  # add a "skill" to the robots skillset the control system will send a string with the ls_item and action and here we will look if we have a matching skill to execute
  # the item_modell defines the patterns which have to be used by the robot on multiple racks and or multiple samples in a rackpattern
  # inner pattern is always dependung on the object that has to be moved and the outer pattern is the pattern for the containers where the objects are stored in.
  # if racks have to be handled it is also an inner pattern cause the object to handle is the rack itself
  # create_item(id=0, ls_item="default", frame=p[0,0,0,0,0,0], actionlist=create_action_list([]), item_model=create_item_model(), lm_id=0, description="default")
  # create_item_model(inner=create_pattern(), outer=create_pattern(), description="default")
  # ITEM_MAP.append(create_item(id=1, ls_item="Home", frame=F1_uLM_Home, actionlist=[ActionManipulator.MOVE_TO], description="uLM Move To Home"))
  # ITEM_MAP.append(create_item(id=2, ls_item="InputStation", frame=F2_uLM_Input, actionlist=[ActionManipulator.PICK, ActionManipulator.PLACE], item_model=create_item_model(inner=Patterns.INPUT), description="uLM Pick and Place samples from Input"))
  # ITEM_MAP.append(create_item(id=3, ls_item="InputCapture", frame=F3_Cap_Input, actionlist=[ActionCamera.INSPECT, ActionManipulator.MOVE_TO], description="uLM Inspect samples from Input and Move To Capture Position"))
  # ITEM_MAP.append(create_item(id=4, ls_item="Bin", frame=F4_uLM_Bin, actionlist=[ActionManipulator.PLACE], description="uLM Place Cap to Bin"))
  # ITEM_MAP.append(create_item(id=5, ls_item="StationaryGripper", frame=F5_uLM_Gripper, actionlist=[ActionManipulator.PICK, ActionManipulator.PLACE, ActionManipulator.DECAP, ActionManipulator.MOVE_TO, ActionManipulator.GRASP, ActionManipulator.RELEASE], description=" uLM stationary gripper"))
  # ITEM_MAP.append(create_item(id=6, ls_item="CobasRack", frame=F6_uLM_Cobas_R, actionlist=[ActionManipulator.PICK, ActionManipulator.PLACE], item_model=create_item_model(outer=Patterns.COBAS_MAGAZINE), description="uLM Cobas Racks Pick and Place"))
  # ITEM_MAP.append(create_item(id=7, ls_item="CobasMagazine", frame=F7_uLM_Coba_Mag, actionlist=[ActionManipulator.PICK, ActionManipulator.PLACE], item_model=create_item_model(inner=Patterns.COBAS, outer=Patterns.COBAS_MAGAZINE), description="uLM Cobas Magazine Samples Pick and Place"))
  # ITEM_MAP.append(create_item(id=8, ls_item="DetectCobasRacks", frame=F8_Cap_Cobas_LM, actionlist=[ActionCamera.DETECT_OBJECTS, ActionManipulator.MOVE_TO], lm_id=2, description="uLM Cobas Rack Detection and Move To Capture"))
  # ITEM_MAP.append(create_item(id=9, ls_item="TaraMagazine", frame=F9_uLM_Tara, actionlist=[ActionManipulator.PICK, ActionManipulator.PLACE], item_model=create_item_model(inner=Patterns.TARA), description="uLM Centrifuge Tara Pick and Place"))
  # ITEM_MAP.append(create_item(id=10, ls_item="CentrifugeCapture", frame=F10_Cap_CF, actionlist=[ActionManipulator.MOVE_TO, ActionCamera.DETECT], lm_id=1, description="Centrifuge Device Move to Capture Pos and Detect Landmarks"))
  # ITEM_MAP.append(create_item(id=11, ls_item="Centrifuge", frame=F11_CF_PiPl, actionlist=[ActionManipulator.PICK, ActionManipulator.PLACE], description="Centrifuge Device Rack Pick and Place"))
  # ITEM_MAP.append(create_item(id=12, ls_item="CentrifugeMagazine", frame=F12_uLM_CF_Mag, actionlist=[ActionManipulator.PICK, ActionManipulator.PLACE], item_model=create_item_model(inner=Patterns.CENTRIFUGE, outer=Patterns.CENTRIFUGE_MAGAZINE), description=" uLM Centrifuge Magazin Pick and Place"))
  # ITEM_MAP.append(create_item(id=13, ls_item="CentrifugeRack", frame=F13_uLM_CF_R, actionlist=[ActionManipulator.PICK, ActionManipulator.PLACE], item_model=create_item_model(outer=Patterns.CENTRIFUGE_MAGAZINE), description="uLM Centrifuge Magazin Pick and Place Racks"))
  # ITEM_MAP.append(create_item(id=14, ls_item="DailyArchive", frame=F14_uLM_Archive, actionlist=[ActionManipulator.PICK, ActionManipulator.PLACE], item_model=create_item_model(inner=Patterns.ARCHIVE), description="uLM Pick and Place samples from Archive Rack"))
  # ITEM_MAP.append(create_item(id=15, ls_item="NokRack", frame=F15_uLM_Nok, actionlist=[ActionManipulator.PICK, ActionManipulator.PLACE], item_model=create_item_model(inner=Patterns.NOK), description="uLM Pick and Place samples from Nok Rack"))
  # ITEM_MAP.append(create_item(id=16, ls_item="CobasInput", frame=F16_Cobas_Input, actionlist=[ActionManipulator.PLACE], description="uLM Place Cobasrack in Cobas Device"))
  # ITEM_MAP.append(create_item(id=17, ls_item="CobasInputCapture", frame=F17_Cobas_Cap, actionlist=[ActionCamera.DETECT, ActionManipulator.MOVE_TO], lm_id=3, description="uLM Place Cobasrack in Cobas Device"))
  # ITEM_MAP.append(create_item(id=18, ls_item="XN550Input", frame=F18_XN550_Input, actionlist=[ActionManipulator.PICK, ActionManipulator.PLACE], item_model=create_item_model(inner=Patterns.SYSMEX_XN550, outer=Patterns.DRAWER_XN550), lm_id=4, description="uLM Pick and Place Samples in or out of XN550 Racks"))
  # ITEM_MAP.append(create_item(id=19, ls_item="XN550Capture", frame=F19_XN550_Cap, actionlist=[ActionCamera.DETECT, ActionManipulator.MOVE_TO], lm_id=4, description="uLM Move To and Capture LM XN550"))
  # ITEM_MAP.append(create_item(id=20, ls_item="XN550Drawer", frame=F20_XN550_Draw, actionlist=[ActionManipulator.DRAWER_OPEN, ActionManipulator.DRAWER_CLOSE], item_model=create_item_model(inner=Patterns.DRAWER_XN550), lm_id=4, description="uLM Open and close Drawer XN550"))
  # ITEM_MAP.append(create_item(id=21, ls_item="XN550Button", frame=F21_XN550_Btn, actionlist=[ActionManipulator.PUSH], lm_id=4, description="uLM Push XN550 Button"))
  # ITEM_MAP.append(create_item(id=22, ls_item="AMR", frame=p[0,0,0,0,0,0], actionlist=[ActionAMR.READ, ActionAMR.LOAD_MISSION, ActionAMR.START_MISSION, ActionAMR.NAVIGATE, ActionAMR.ACKNOWLEDGE], description="all AMR actions"))



  # ITEM_MAP.append(create_item(id=31, ls_item="TestLM", frame=TestLM, actionlist=[ActionManipulator.PICK, ActionManipulator.PLACE], item_model=create_item_model(inner=Rack.SYSMEX_CS2500), lm_id=5, description="LM Test"))
  # Fills the Vision Config List with Projectrelated Data
  # workspaceid and skillid are highly robominds related so probably will not stay like this in the future
  # sample detection: dx and dy are used to calculate the positions in a rack and given by the offset which will be applied in order to assign the sample to a place in the rack
  # create_vision_config(workspace_id="", skill_id="", item_id=-1, capture_pos=p[0,0,0,0,0,0], dx=0, dy=0, target_origin=p[0,0,0,0,0,0], selector="default", description="default")
  # VISION_CONFIG_MAP.append(create_vision_config(workspace_id="96017791-f581-4e9e-93da-6951695fccc8", skill_id="8885cfe1-6784-4293-bd26-52ebdc67bf95", capture_pos=F10_Cap_CF, target_origin=p[0,0,0,0,0,0], item_id=11, description="LM Detect CF"))
  # VISION_CONFIG_MAP.append(create_vision_config(workspace_id="96017791-f581-4e9e-93da-6951695fccc8", skill_id="8885cfe1-6784-4293-bd26-52ebdc67bf95", capture_pos=F8_Cap_Cobas_LM, target_origin=p[0,0,0,0,0,0], item_id=8, description="LM Detect Cobas Racks"))
  # VISION_CONFIG_MAP.append(create_vision_config(workspace_id="8f0ad01c-dc36-4fdd-b295-0b6b4a38b89a", skill_id="afdc9e13-ea83-40d6-a805-bb041453d2e5", capture_pos=F3_Cap_Input, target_origin=F2_uLM_Input, item_id=3, description="Lab Solution Input Capture"))
  # VISION_CONFIG_MAP.append(create_vision_config(workspace_id="96017791-f581-4e9e-93da-6951695fccc8", skill_id="8885cfe1-6784-4293-bd26-52ebdc67bf95", capture_pos=F19_XN550_Cap, target_origin=F18_XN550_Input, item_id=18, description="Input XN550"))
  # VISION_CONFIG_MAP.append(create_vision_config(workspace_id="96017791-f581-4e9e-93da-6951695fccc8", skill_id="8885cfe1-6784-4293-bd26-52ebdc67bf95", capture_pos=F19_XN550_Cap, target_origin=POS_Z, item_id=19, description="LM Detect XN550F"))
  # VISION_CONFIG_MAP.append(create_vision_config(workspace_id="96017791-f581-4e9e-93da-6951695fccc8", skill_id="8885cfe1-6784-4293-bd26-52ebdc67bf95", capture_pos=F10_Cap_CF, target_origin=POS_Z, item_id=10, description="LM Detect CF"))
  # VISION_CONFIG_MAP.append(create_vision_config(workspace_id="96017791-f581-4e9e-93da-6951695fccc8", skill_id="8885cfe1-6784-4293-bd26-52ebdc67bf95", capture_pos=F19_XN550_Cap, target_origin=F20_XN550_Draw, item_id=20, description="Drawer XN550"))
  # VISION_CONFIG_MAP.append(create_vision_config(workspace_id="96017791-f581-4e9e-93da-6951695fccc8", skill_id="8885cfe1-6784-4293-bd26-52ebdc67bf95", capture_pos=F19_XN550_Cap, target_origin=F21_XN550_Btn, item_id=21, description="Button XN550"))
  # VISION_CONFIG_MAP.append(create_vision_config(workspace_id="96017791-f581-4e9e-93da-6951695fccc8", skill_id="8885cfe1-6784-4293-bd26-52ebdc67bf95", capture_pos=TestLMCap, target_origin=p[0,0,0,0,0,0], item_id=30, description="Button XN550"))
  # VISION_CONFIG_MAP.append(create_vision_config(workspace_id="96017791-f581-4e9e-93da-6951695fccc8", skill_id="8885cfe1-6784-4293-bd26-52ebdc67bf95", capture_pos=TestLMCap, target_origin=TestLM, item_id=31, description="Button XN550"))

  # VISION_CONFIG_MAP.append(create_vision_config(workspace_id="96017791-f581-4e9e-93da-6951695fccc8", skill_id="8885cfe1-6784-4293-bd26-52ebdc67bf95", target_origin=p[0,0,0,0,0,0], item_id=11, description="LM Detect CF"))
  # VISION_CONFIG_MAP.append(create_vision_config(workspace_id="96017791-f581-4e9e-93da-6951695fccc8", skill_id="8885cfe1-6784-4293-bd26-52ebdc67bf95", target_origin=p[0,0,0,0,0,0], item_id=8, description="LM Detect Cobas Racks"))
  # VISION_CONFIG_MAP.append(create_vision_config(workspace_id="8f0ad01c-dc36-4fdd-b295-0b6b4a38b89a", skill_id="afdc9e13-ea83-40d6-a805-bb041453d2e5", target_origin=F2_uLM_Input, item_id=3, description="Lab Solution Input Capture"))
  # VISION_CONFIG_MAP.append(create_vision_config(workspace_id="96017791-f581-4e9e-93da-6951695fccc8", skill_id="8885cfe1-6784-4293-bd26-52ebdc67bf95", target_origin=F18_XN550_Input, item_id=18, description="Input XN550"))
  # VISION_CONFIG_MAP.append(create_vision_config(workspace_id="96017791-f581-4e9e-93da-6951695fccc8", skill_id="8885cfe1-6784-4293-bd26-52ebdc67bf95", target_origin=POS_Z, item_id=19, description="LM Detect XN550F"))
  # VISION_CONFIG_MAP.append(create_vision_config(workspace_id="96017791-f581-4e9e-93da-6951695fccc8", skill_id="8885cfe1-6784-4293-bd26-52ebdc67bf95", target_origin=POS_Z, item_id=10, description="LM Detect CF"))
  # VISION_CONFIG_MAP.append(create_vision_config(workspace_id="96017791-f581-4e9e-93da-6951695fccc8", skill_id="8885cfe1-6784-4293-bd26-52ebdc67bf95", target_origin=F20_XN550_Draw, item_id=20, description="Drawer XN550"))
  # VISION_CONFIG_MAP.append(create_vision_config(workspace_id="96017791-f581-4e9e-93da-6951695fccc8", skill_id="8885cfe1-6784-4293-bd26-52ebdc67bf95", target_origin=F21_XN550_Btn, item_id=21, description="Button XN550"))
  # VISION_CONFIG_MAP.append(create_vision_config(workspace_id="96017791-f581-4e9e-93da-6951695fccc8", skill_id="8885cfe1-6784-4293-bd26-52ebdc67bf95", target_origin=p[0,0,0,0,0,0], item_id=30, description="Button XN550"))
  # VISION_CONFIG_MAP.append(create_vision_config(workspace_id="96017791-f581-4e9e-93da-6951695fccc8", skill_id="8885cfe1-6784-4293-bd26-52ebdc67bf95", target_origin=TestLM, item_id=31, description="Button XN550"))

  # local inputrack = find_pattern_by_name("INPUT")
  # INSPECT_CONFIG_MAP.append(create_inspect_config(item_id=3, dx=inputrack.pattern_width[0]/(inputrack.pattern_size[0]-1), dy=inputrack.pattern_width[1]/(inputrack.pattern_size[1]-1), rack_size=inputrack.pattern_size , description="Input Capture"))
  # # Fills the Landmark List with Projectrelated Data
  # # create_landmark(lm_id=0, marker_id=-1, marker_size=0.1, marker_type="aruco_7x7", capture_pos=p[0,0,0,0,0,0], init_frame=p[0,0,0,0,0,0], search_offset=[0,0,0], actual_frame=p[0,0,0,0,0,0], description="")
  # LANDMARK_MAP.append(create_landmark(lm_id=1, marker_id=3, marker_size=0.1, marker_type="aruco_7x7", capture_pos = F10_Cap_CF, init_frame=p[-0.617789, -0.065471, 0.07918, 0.020983, -0.012695, 1.512066], search_offset=[0.15, 0.15, 0.1], actual_frame=p[-0.617789, -0.065471, 0.07918, 0.020983, -0.012695, 1.512066], description="LM CF Lid"))
  # LANDMARK_MAP.append(create_landmark(lm_id=2, marker_id=-1, marker_size=0.0085, marker_type="aruco_4x4", capture_pos = F8_Cap_Cobas_LM, init_frame=p[0,0,0,0,0,0], search_offset=[0.15, 0.15, 0.1], actual_frame=POS_Z, description="LM Cobas Rack Detection"))
  # LANDMARK_MAP.append(create_landmark(lm_id=3, marker_id=0, marker_size=0.1, marker_type="aruco_7x7", capture_pos = F17_Cobas_Cap, init_frame=p[-0.667,-0.194,0.100,0,0,0], search_offset=[0.15, 0.15, 0.1], actual_frame=POS_Z, description="LM Cobas Cap"))
  # LANDMARK_MAP.append(create_landmark(lm_id=4, marker_id=4, marker_size=0.1, marker_type="aruco_7x7", capture_pos = F19_XN550_Cap, init_frame=p[0.124,-0.976,0.355,-0.008,0.025,3.131], search_offset=[0.15, 0.15, 0.1], actual_frame=p[0,0,0,0,0,0], description="LM XN550 Cap"))
  # LANDMARK_MAP.append(create_landmark(lm_id=5, marker_id=0, marker_size=0.1, marker_type="aruco_7x7", capture_pos = TestLMCap, init_frame=p[-0.49,-0.144,0.092,0,-0.008,0.001], search_offset=[0.15, 0.15, 0.1], actual_frame=POS_Z, description="LM Test"))
  # # Configuration of all movement related parameters
  # # create_movement(id=0, hh_approach=POS_Z, h_approach=POS_Z, approach=POS_Z, h_target=POS_Z, target=POS_Z, retract=POS_Z, h_retract=POS_Z, hh_retract=POS_Z, h_frame=POS_Z, frame=POS_Z, speed=1, acceleration=1, description="default")
  # MOVEMENT_MAP.append(create_movement(description="TestLMCap", frame=TestLMCap, actionlist=[ActionManipulator.MOVE_TO]))
  # MOVEMENT_MAP.append(create_movement(description="TestLM", frame=TestLM, actionlist=[ActionManipulator.PICK,ActionManipulator.PLACE],
  #         approach=p[0,0,0.1,0,0,0],
  #         retract=p[0,0,0.1,0,0,0]))
  # MOVEMENT_MAP.append(create_movement(description="Home - MOVE_TO", frame=F1_uLM_Home, actionlist=[ActionManipulator.MOVE_TO]))
  # MOVEMENT_MAP.append(create_movement(description="Input - PICK&PLACE", frame=F2_uLM_Input, actionlist=[ActionManipulator.PICK,ActionManipulator.PLACE],
  #         approach=p[0,0,0.1,0,0,0],
  #         retract=p[0,0,0.1,0,0,0]))
  # MOVEMENT_MAP.append(create_movement(description="Capture Input - MOVE_TO", frame=F3_Cap_Input, actionlist=[ActionManipulator.MOVE_TO]))
  # MOVEMENT_MAP.append(create_movement(description="BIN - PLACE", frame=F4_uLM_Bin, actionlist=[ActionManipulator.PLACE],
  #         approach=p[0,0,0.1,0,0,0],
  #         retract=p[0,0,0.1,0,0,0]))
  # MOVEMENT_MAP.append(create_movement(description="Gripper - Move To", frame=F5_uLM_Gripper, actionlist=[ActionManipulator.MOVE_TO],
  #         approach=p[0,0,0.1,0,0,0]))
  # MOVEMENT_MAP.append(create_movement(description="Gripper - Pick", frame=F5_uLM_Gripper, actionlist=[ActionManipulator.PICK],
  #         retract=p[0,0,0.1,0,0,0]))
  # MOVEMENT_MAP.append(create_movement(description="Gripper - Place", frame=F5_uLM_Gripper, actionlist=[ActionManipulator.PLACE],
  #         approach=p[0,0,0.1,0,0,0]))
  # MOVEMENT_MAP.append(create_movement(description="CobasRack Pick & Place", frame=F6_uLM_Cobas_R, actionlist=[ActionManipulator.PICK,ActionManipulator.PLACE],
  #         approach=p[0,0,0.1,0,0,0],
  #         target=p[0,0,0,0,0,d2r(90)],
  #         retract=p[0,0,0.1,0,0,0]))
  # MOVEMENT_MAP.append(create_movement(description="CobasMagazine Pick & Place", frame=F7_uLM_Coba_Mag, actionlist=[ActionManipulator.PICK,ActionManipulator.PLACE],
  #         approach=p[0,0,0.1,0,0,0],
  #         target=p[0,0,0,0,0,-d2r(90)],
  #         retract=p[0,0,0.1,0,0,0]))
  # MOVEMENT_MAP.append(create_movement(description="Capture Position Cobas Landmarks", frame=F8_Cap_Cobas_LM, actionlist=[ActionManipulator.MOVE_TO]))
  # MOVEMENT_MAP.append(create_movement(description="TaraMagazine - PICK & PLACE", frame=F9_uLM_Tara, actionlist=[ActionManipulator.PICK,ActionManipulator.PLACE],
  #         approach=p[0,0,0.13,0,0,0],
  #         target=p[0,0,0,0,0,-d2r(90)],
  #         retract=p[0,0,0.13,0,0,0]))
  # MOVEMENT_MAP.append(create_movement(description="Capture Position - Centrifuge LM", frame=F10_Cap_CF,actionlist=[ActionManipulator.MOVE_TO]))
  # MOVEMENT_MAP.append(create_movement(description="Pick and Place Racks - Centrifuge Lid", frame=F11_CF_PiPl, actionlist=[ActionManipulator.PICK,ActionManipulator.PLACE],
  #         approach=p[0,0,0.3,0,0,0],
  #         retract=p[0,0,0.3,0,0,0]))
  # MOVEMENT_MAP.append(create_movement(description="Pick and Place Samples - Centrifuge on uLM", frame=F12_uLM_CF_Mag, actionlist=[ActionManipulator.PICK,ActionManipulator.PLACE],
  #         approach=p[0,0,0.13,0,0,0],
  #         retract=p[0,0,0.13,0,0,0]
  #         ))
  # MOVEMENT_MAP.append(create_movement(description="Pick and Place Racks - Centrifuge on uLM", frame=F13_uLM_CF_R, actionlist=[ActionManipulator.PICK,ActionManipulator.PLACE],
  #         approach=p[0,0,0.15,0,0,0],
  #         retract=p[0,0,0.15,0,0,0]
  #         ))

  # MOVEMENT_MAP.append(create_movement(description="Pick and Place Samples XN550 Racks in Device", frame=F18_XN550_Input, actionlist=[ActionManipulator.PICK,ActionManipulator.PLACE],
  #         approach=p[0,0,0.1,0,0,0],
  #         target = p[0,0,0,0,0,d2r(90)],
  #         retract=p[0,0,0.1,0,0,0]
  #         ))
  # MOVEMENT_MAP.append(create_movement(description="Capture LM XN550", frame=F19_XN550_Cap, actionlist=[ActionManipulator.MOVE_TO]))
  # MOVEMENT_MAP.append(create_movement(description="Open XN550 Drawer ", frame=F20_XN550_Draw, actionlist=[ActionManipulator.DRAWER_OPEN],
  #         h_approach=p[0.07,0,0.1,0,0,0],
  #         approach=p[0,0,0.1,0,0,0],
  #         target = p[0,0,0,0,0,d2r(90)],
  #         retract=p[0.07,0,0,0,0,0],
  #         h_retract=p[0.07,0,0.1,0,0,0]
  #         ))
  # MOVEMENT_MAP.append(create_movement(description="Close XN550 Drawer ", frame=F20_XN550_Draw, actionlist=[ActionManipulator.DRAWER_CLOSE],
  #         h_approach=p[0.07,0,0.1,0,0,0],
  #         approach=p[0.07,0,0,0,0,0],
  #         target = p[0,0,0,0,0,d2r(90)],
  #         retract=p[0,0,0.1,0,0,0],
  #         h_retract=p[0.07,0,0.1,0,0,0]
  #         ))
  # MOVEMENT_MAP.append(create_movement(description="Push XN550 Button ", frame=F21_XN550_Btn, actionlist=[ActionManipulator.PUSH],
  #         approach=p[0,0,0.15,0,0,0],
  #         retract=p[0,0,0.15,0,0,0]
  #         ))
  # MOVEMENT_MAP.append(create_movement(description="Capture Position 2 Input", frame=F_Cap_Input2,actionlist=[ActionManipulator.MOVE_TO]))



  $ 19 "Script: SCRIPT Objects V0.1.script"
  #*****************************************************
  # customer          :   INTERNAL
  # project name      :
  #****************************************************
  # controller        :   UR
  # software          :   5.17.3
  #****************************************************
  # author            :   P. Koehnke
  # Copyright (c)     :   United Robotics Group
  #                       An der Riede 2
  #                       28816 Stuhr
  #                       Germany
  #****************************************************
  # description       :   object database
  # version:      	:   0.1
  # created           :   09.10.2024
  # updated           :
  #****************************************************
  # modifications     :
  #
  # date              :
  # name              :
  # reason            :
  #****************************************************

  def create_object_2(id=0, name="", type=0, dimension=struct(length=0, width=0, height=0, diameter=0), gripper_offset=p[0,0,0,0,0,0]):
      return struct(id=id, name=name, type=type, dimension=dimension, gripper_offset=gripper_offset)
  end

  OBJ = create_object_2()
  OBJs = make_list(0, create_object_2(), 50)

  OBJs.append(create_object_2(id=1, name="rack centrifuge", type=1, dimension=struct(length=0, width=0, height=0.106, diameter=0.020), gripper_offset=p[0,0,0.095,0,0,2.356]))
  OBJs.append(create_object_2(id=2, name="sample tube 1", type=2, dimension=struct(length=0, width=0, height=0.106, diameter=0.015), gripper_offset=p[0,0,0,0,0,0]))
  OBJs.append(create_object_2(id=3, name="rack sarstedt", type=3, dimension=struct(length=0, width=0, height=0.100, diameter=0.020), gripper_offset=p[0,0,0,0,0,0]))
  OBJs.append(create_object_2(id=4, name="Lab bottle", type=4, dimension=struct(length=0, width=0, height=0.100, diameter=0.030), gripper_offset=p[0,0,0.2,0,0,0]))
  OBJs.append(create_object_2(id=5, name="Vial", type=5, dimension=struct(length=0, width=0, height=0.100, diameter=0.0275), gripper_offset=p[0,0,0,0,0,0]))
  OBJs.append(create_object_2(id=6, name="Container", type=6, dimension=struct(length=0.0, width=0.0, height=0, diameter=0.0), gripper_offset=p[0,0,0,0,0,0]))
  OBJs.append(create_object_2(id=7, name="Target_container", type=7, dimension=struct(length=0.06, width=0.06, height=0.134, diameter=0.05), gripper_offset=p[0,0,0,0,0,0]))
  OBJs.append(create_object_2(id=8, name="Spatula", type=8, dimension=struct(length=0.03, width=0.03, height=0.23, diameter=0.05), gripper_offset=p[0,0,0,0,0,0]))
  OBJs.append(create_object_2(id=9, name="rack pipet", type=9, dimension=struct(length=0.03, width=0.03, height=0.23, diameter=0.05), gripper_offset=p[0,0,0,0,0,0]))

  def create_jig_2(id=0, name="", type=0, capacity=0, jig_offset=p[0,0,0,0,0,0]):
      # iformation about used jigs
      return struct(id=id, name=name, type=type, capacity=capacity, jig_offset=jig_offset)
  end

  JIG2 = create_jig_2()
  JIGs = make_list(0, create_jig_2(), 20)

  JIGs.append(create_jig_2(id=1, name="3FG", type=1, capacity=1, jig_offset=p[0,0,0,0,0,0]))
  JIGs.append(create_jig_2(id=2, name="jig input", type=2, capacity=1, jig_offset=p[0,0,0,0,0,-3.927]))
  JIGs.append(create_jig_2(id=3, name="jig output", type=3, capacity=1, jig_offset=p[0,0,0,0,0,0.78]))
  JIGs.append(create_jig_2(id=6, name="jig bin", type=6, capacity=1, jig_offset=p[0,0,0,0,0,0]))
  JIGs.append(create_jig_2(id=7, name="jig sarstedt racks", type=7, capacity=1, jig_offset=p[0,0,-0.02,0,0,0]))
  JIGs.append(create_jig_2(id=8, name="NoK Bin", type=8, capacity=1, jig_offset=p[0,0,0,0,0,0]))
  JIGs.append(create_jig_2(id=9, name="Pick bott jig", type=9, capacity=1, jig_offset=p[0,0,0,0,0,0]))
  JIGs.append(create_jig_2(id=10, name="Place bott jig", type=10, capacity=1, jig_offset=p[0,0,0,0,0,0]))
  JIGs.append(create_jig_2(id=11, name="bottle shake jig", type=11, capacity=1, jig_offset=p[0,0,0,0,0,0]))
  JIGs.append(create_jig_2(id=12, name="Pick Vial jig", type=12, capacity=1, jig_offset=p[0,0,0,0,0,0]))
  JIGs.append(create_jig_2(id=13, name="Place Vial jig", type=13, capacity=1, jig_offset=p[0,0,0,0,0,0]))
  JIGs.append(create_jig_2(id=14, name="Liquid transfer jig", type=14, capacity=1, jig_offset=p[0,0,0,0,0,0]))
  JIGs.append(create_jig_2(id=15, name="Pick station jig", type=15, capacity=1, jig_offset=p[0,0,0,0,0,0]))
  JIGs.append(create_jig_2(id=16, name="Place station jig", type=16, capacity=1, jig_offset=p[0,0,0,0,0,0]))
  JIGs.append(create_jig_2(id=17, name="Weigh station jig", type=17, capacity=1, jig_offset=p[0,0,0,0,0,0]))
  JIGs.append(create_jig_2(id=18, name="Pick station 1", type=18, capacity=1, jig_offset=p[0,0,0,0,0,0]))
  JIGs.append(create_jig_2(id=19, name="Pick station 2", type=19, capacity=1, jig_offset=p[0,0,0,0,0,0]))
  JIGs.append(create_jig_2(id=20, name="Pick station 3", type=20, capacity=1, jig_offset=p[0,0,0,0,0,0]))
  JIGs.append(create_jig_2(id=21, name="Tilt station jig", type=21, capacity=1, jig_offset=p[0,0,0,0,0,0]))
  JIGs.append(create_jig_2(id=22, name="Swab station jig", type=22, capacity=1, jig_offset=p[0,0,0,0,0,0]))
  $ 20 "Script: Powder_all_newspats.script"
  #global SERVER_IP   = "192.168.12.139"


  global tcp_dosing = p[0,0,0.15052,3.1415,0,0]
  global tcp_default = p[0,0,0.161,3.1415,0,0]

  global container_id = 0
  global powder_id  = 0
  global bulk_density = 0
  global H          = 0
  global H_c          = 0
  global mouth_d     = 0
  global mouth_sh    = 0
  global length_c     = 0
  global diameter   = 0
  global empty_weight_g  = 0
  global volume_ml    = 0
  global shape_code   = 0
  global flow_code   = 0
  global shape = ""
  global Flowability = ""
  global full_weight_g = 0
  global cent_edge = 0
  global pick_2_base = 0.2 # distance from tcp to base of picking table
  global wall_thickness = 0.002

  def read_db_data():

    socket_open(SERVER_IP, SERVER_PORT)
    sleep(0.5)
    socket_send_string("GET_DATACODE_FLOATS")
    sleep(5)

    local fl = socket_read_ascii_float(14)
    socket_close()

    global container_id = fl[1]
    global powder_id = fl[2]
    global bulk_density = fl[3]
    global H          = fl[4]/1000
    global H_c          = fl[5]/1000
    global mouth_d     = fl[6]/1000
    global mouth_sh    = fl[7]/1000
    global length_c     = fl[8]/1000
    global diameter   = fl[9]/1000
    global empty_weight_g = fl[10]
    global volume_ml    = fl[11]
    global full_weight_g = fl[12]
    global flow_code   = fl[13]
    global shape_code   = fl[14]

  	if (flow_code == 1.0):
  		global Flowability = "MEDIUM"
  	elif (flow_code == 2.0):
  		global Flowability = "LOW"
  	else:
  		global Flowability = "HIGH"
  	end

  	if ( shape_code == 1.0):
  		shape = "cylindrical"
  		cent_edge =  diameter
  	else:
  		shape = "cubical"
  		cent_edge =  length_c
  	end

  	read_spatula_data()

  end

  def send_picking_info(Pow_name, target_weight):
    socket_open(SERVER_IP, SERVER_PORT)
    cmd = "PICK:"+Pow_name+";"+to_str(target_weight)
    socket_send_string(cmd)
    sleep(0.1)
    socket_close()
  end

  #### POTS ####
  def tilt_send(angle):
  	socket_open(SERVER_IP, SERVER_PORT)
  	angle = 92.0 - angle
  	socket_send_string("TILT:"+to_str(angle))
  	sync()
  	sleep(0.5)
  	socket_close()
  end

  def CW_Rotate(angle):
  	socket_open(SERVER_IP, SERVER_PORT)
  	socket_send_string("CWROTATE:"+to_str(angle))
  	sync()
  	sleep(0.5)
  	socket_close()
  end

  def CCW_Rotate(angle):
  	socket_open(SERVER_IP, SERVER_PORT)
  	socket_send_string("CCWROTATE:"+to_str(angle))
  	sync()
  	sleep(0.5)
  	socket_close()
  end

  def CW_full_Rotate():
  	socket_open(SERVER_IP, SERVER_PORT)
  	socket_send_string("FULLROTATE:"+to_str(1))
  	sync()
  	sleep(0.5)
  	socket_close()
  end

  def CCW_full_Rotate():
  	socket_open(SERVER_IP, SERVER_PORT)
  	socket_send_string("FULLROTATE:"+to_str(-1))
  	sync()
  	sleep(0.5)
  	socket_close()
  end

  def tilt_to_home():
  	socket_open(SERVER_IP, SERVER_PORT)
  	socket_send_string("HOME")
  	sync()
  	sleep(0.5)
  	socket_close()
  end
  #######
  def vibration_1():
  	set_analog_out(0,0.4)
  	sleep(1)
  	set_analog_out(0,0.0)
  	sleep(0)
  end

  def vibration_2():
  	set_analog_out(0,0.4)
  	sleep(0.8)
  	set_analog_out(0,0.0)
  	sleep(0.2)
  end

  def vibration_3():
  	set_analog_out(0,0.4)
  	sleep(0.5)
  	set_analog_out(0,0.0)
  	sleep(0.3)
  end

  def vibration_4():
  	set_analog_out(0,0.4)
  	sleep(0.5)
  	set_analog_out(0, 0.0)
  	sleep(0.5)
  end

  def vibration_5():
  	set_analog_out(0,0.4)
  	sleep(0.2)
  	set_analog_out(0, 0.0)
  	sleep(0.8)
  end

  ##################

  global gear_2_holder = 0.018
  global hinge_2_base = 0.0421
  global TCP_2_tip_x = 0.0047
  global spatula_len = 0.182
  global spatula_offset = p[TCP_2_tip_x,0,spatula_len,0,0,0]
  global SPATULA_L_VOL_ML = 0.0
  global SPATULA_M_VOL_ML = 0.0
  global SPATULA_S_VOL_ML = 0.0
  global SPATULA_FLAT_M_VOL_ML  = 0.0
  global SPATULA_FLAT_S_VOL_ML  = 0.0

  global DB_SPATULA_L_DEPTH = 0.0
  global DB_SPATULA_M_DEPTH = 0.0
  global DB_SPATULA_S_DEPTH = 0.0
  global DB_SPATULA_FLAT_M_DEPTH = 0.0
  global DB_SPATULA_FLAT_S_DEPTH = 0.0
  global DB_SPATULA_L_MID = 0.0
  global DB_SPATULA_M_MID = 0.0
  global DB_SPATULA_S_MID = 0.0
  global DB_SPATULA_FLAT_M_MID = 0.0
  global DB_SPATULA_FLAT_S_MID = 0.0
  global DB_SPATULA_L_RY = 0.0
  global DB_SPATULA_M_RY = 0.0
  global DB_SPATULA_S_RY = 0.0
  global DB_SPATULA_FLAT_M_RY = 0.0
  global DB_SPATULA_FLAT_S_RY = 0.0

  def read_spatula_data():
  	socket_open(SERVER_IP, SERVER_PORT)
  	sleep(0.2)
  	socket_send_string("GET_SPATULA_FLOATS")
  	sleep(0.5)
  	local fl = socket_read_ascii_float(25)
  	socket_close()

  	global DB_SPATULA_L_DEPTH = fl[1]/1000
  	global DB_SPATULA_L_MID = fl[2]/2000
  	global SPATULA_L_VOL_ML = fl[3]
  	global DB_SPATULA_L_RY = fl[4]
  	global DB_SPATULA_M_DEPTH = fl[6]/1000
  	global DB_SPATULA_M_MID = fl[7]/2000
  	global SPATULA_M_VOL_ML = fl[8]
  	global DB_SPATULA_M_RY = fl[9]
  	global DB_SPATULA_S_DEPTH = fl[11]/1000
  	global DB_SPATULA_S_MID = fl[12]/2000
  	global SPATULA_S_VOL_ML = fl[13]
  	global DB_SPATULA_S_RY = fl[14]
  	global DB_SPATULA_FLAT_M_DEPTH = fl[16]/1000
  	global DB_SPATULA_FLAT_M_MID = fl[17]/2000
  	global SPATULA_FLAT_M_VOL_ML = fl[18]
  	global DB_SPATULA_FLAT_M_RY = fl[19]
  	global DB_SPATULA_FLAT_S_DEPTH = fl[21]/1000
  	global DB_SPATULA_FLAT_S_MID = fl[22]/2000
  	global SPATULA_FLAT_S_VOL_ML = fl[23]
  	global DB_SPATULA_FLAT_S_RY = fl[24]
  end

  def correction_reset():
  	global g_k = 0.0
  	global g_depth_corr = 0.0
  	global g_prev_cum_w = weight_value
  end

  def params_init():

  	global scoop_status= ""
  	global w_dosed_total = 0.0
  	global last_scale = 0.0
  	global tilt_angle_sent = 0.0
  	global level = 0.0
  	global target_g = 0.0
  	global angle_max = 65
  	global angle_min = 30
  	global gain_per_percent = (angle_max - angle_min)/100
  	global ry_deg_safe = 0
  	global ry_deg = 0
  	global delta_count=0

  	global scoop_ct = 0
  	global error_sum = 0.0
  	global error_sq_sum = 0.0
  	global scoop_g = 0.0

  	global g_k =0.0
  	global g_eta = 0.3

  	global g_gain_scale = 0.07
  	global g_k_min = 0.0
  	global g_k_max = 0.09

  	# ---------- Damping ----------
  	global g_alpha_under = 0.75   # aggressive when undershooting
  	global g_alpha_over  = 0.60   # conservative when overshooting

  	# ---------- Search ----------
  	global g_engagement_min = 0.05
  	global g_search_step = 0.01      # 3 mm

  	# ---------- Deadband ----------
  	global g_tol = 0.02               # 20 mg minimum
  	global g_tol_ratio = 0.05         # ±5% of target

  	# ---------- Limits ----------
  	global g_corr_max = 0.020         # 20 mm maximum correction

  	# ---------- States ----------
  	global g_depth_corr = 0.0
  	global g_prev_cum_w = -1.0
  	global z_ratio = 0.0
  	global z_offset = 0.0
  end

  def clamp(x, lo, hi):
  	if(x<lo):
  		return lo
  	elif (x>hi):
  		return hi
  	else:
  		return x
  	end
  end

  def compute_level_percent(W_now, weight_value):   # W_now = container+powder, weight_value = live scale reading
      global delta = weight_value - last_scale

      if (delta < 0.0):
          delta = 0.0
      end

      global w_dosed_total = w_dosed_total + delta
      global last_scale = weight_value     # update the last scale reading

      local W_eff = W_now - w_dosed_total
      if (W_eff <  empty_weight_g):
          W_eff =  empty_weight_g
      end

      # Compute powder level %
      level = 100.0 * (W_eff -  empty_weight_g) / (full_weight_g -  empty_weight_g)

      # Clamp to 0–100
      level = clamp(level, 0, 100)
    textmsg("deb 1 = ", level)
      return level
  end

  def deg2rad(d):
  	return d*3.141592/180
  end

  def my_abs(val):
  	if (val<0):
  		return -val
  	else:
  		return val
  	end
  end

  def compute_tilt_deg(level_percent):
  	angle = angle_min + gain_per_percent*(100.0-level_percent)

    	textmsg("deb 2 = ", angle)
  	return clamp(angle, angle_min, angle_max)
  end

  def tilt(level_percentage):
  	new_angle = compute_tilt_deg(level_percentage)
    	textmsg("deb angle 1 = ", new_angle)
  	global angle_rel = new_angle - tilt_angle_sent
    	textmsg("deb 2 = ", angle_rel)

  	if my_abs(angle_rel)>2.0:
    		textmsg("deb loop")
  		tilt_send(new_angle)
  		global angle_deg = new_angle
    		textmsg("deb 2 = ", angle_deg)
  		global tilt_angle_sent = new_angle
  		global p_center_vertical = center_pose()
  		global p_center = updated_center_pose(p_center_vertical, angle_deg)
  	end
    	textmsg("deb loop exit")

  	tilt_send(angle_deg)
    	textmsg("deb angle 2 =", angle_deg)

  end

  def compute_scoop_depth(level, weight_value, target_g):

      global scoop_depth_rel = ((100.0-level)/100.0)*(H-mouth_sh)

      if (g_prev_cum_w < 0):
          g_prev_cum_w = weight_value
          g_depth_corr = 0.0

      else:
          global scoop_g = weight_value - g_prev_cum_w
          g_prev_cum_w = weight_value

          local error = target_g - scoop_g
          local engagement = scoop_g / target_g

          local tol = g_tol_ratio * target_g
          if (tol < g_tol):
              tol = g_tol
          end
          if ((engagement < g_engagement_min) and (scoop_g < target_g)):
              g_depth_corr = g_depth_corr + g_search_step
          elif (my_abs(error) <= tol):
  			sync()
          else:
              local error_norm = my_abs(error / target_g)
              local g_target = clamp(g_gain_scale * error_norm,g_k_min,g_k_max)

              g_k = (1.0-g_eta) * g_k + g_eta * g_target
              if (error > 0):
                  local corr = g_k * error
                  g_depth_corr = g_depth_corr +g_alpha_under * corr
              else:
                  local corr = g_k * error
                  g_depth_corr = g_depth_corr +g_alpha_over * corr

              end
              g_depth_corr = clamp(g_depth_corr,-g_corr_max,g_corr_max)

          end
      end
      scoop_depth = scoop_depth_rel + g_depth_corr
      scoop_depth = clamp(scoop_depth, 0.0, H)
      return scoop_depth

  end

  def get_scoop_weight(spatula, bulk_density):

  	local vol = 0

  	if (spatula == "spatula_L"):
  		vol = SPATULA_L_VOL_ML
  		global spatula_depth = DB_SPATULA_L_DEPTH
  		global spatula_mid   = DB_SPATULA_L_MID
  		global spatula_ry    = DB_SPATULA_L_RY

  	elif (spatula == "spatula_M"):
  		vol = SPATULA_M_VOL_ML
  		global spatula_depth = DB_SPATULA_M_DEPTH
  		global spatula_mid   = DB_SPATULA_M_MID
  		global spatula_ry    = DB_SPATULA_M_RY

  	elif (spatula == "spatula_S"):
  		vol = SPATULA_S_VOL_ML
  		global spatula_depth = DB_SPATULA_S_DEPTH
  		global spatula_mid   = DB_SPATULA_S_MID
  		global spatula_ry    = DB_SPATULA_S_RY

  	elif (spatula == "spatula_flat_M"):
  		vol = SPATULA_FLAT_M_VOL_ML
  		global spatula_depth = DB_SPATULA_FLAT_M_DEPTH
  		global spatula_mid   = DB_SPATULA_FLAT_M_MID
  		global spatula_ry    = DB_SPATULA_FLAT_M_RY

  	elif (spatula == "spatula_flat_S"):
  		vol = SPATULA_FLAT_S_VOL_ML
  		global spatula_depth = DB_SPATULA_FLAT_S_DEPTH
  		global spatula_mid   = DB_SPATULA_FLAT_S_MID
  		global spatula_ry    = DB_SPATULA_FLAT_S_RY
  	else:
  		textmsg("Unknown spatula type")
  		return 0.0
  	end
  	global target_g = vol * bulk_density
  	return target_g

  end

  def select_spatula(Flowability, level, diff, bulk_density, mouth_d ):

      local k = 1.1
      global powder_height = (H  - mouth_sh ) * level/100

      if (Flowability == "LOW"):
          local gFM = get_scoop_weight("spatula_flat_M", bulk_density)
  		local mouth_ok_FM = (mouth_d >= 0.05)
  		local level_ok_FM = (spatula_mid  < powder_height)
          local diff_ok_FM  = (diff > k * gFM)
  		local flatM_ok = mouth_ok_FM and level_ok_FM and diff_ok_FM
          if (flatM_ok):
              return "spatula_flat_M"
          else:
              return "spatula_flat_S"
          end
      end

      local gL = get_scoop_weight("spatula_L", bulk_density)
      local mouth_ok_L = (mouth_d  >= 0.05)
      local level_ok_L = (spatula_mid < powder_height)
      local diff_ok_L  = (diff > k * gL)

      local large_ok = mouth_ok_L and level_ok_L and diff_ok_L
      local gM = get_scoop_weight("spatula_M", bulk_density)
      local level_ok_M = (spatula_mid < powder_height)
      local diff_ok_M  = (diff > k * gM)

      local medium_ok = level_ok_M and diff_ok_M

      if (large_ok):
          return "spatula_L"
      elif (medium_ok):
          return "spatula_M"
      else:
          return "spatula_S"
      end
  end

  def after_scoop():
  	set_tcp(tcp_dosing)
  	set_analog_out(0,0.0)
  	tilt_send(angle_deg)
  	sleep(0.5)
  	movel(lifted_pose, a=0.05, v=0.2)
  	movel(move_inside_spill, a=0.05, v=0.2)
  	set_analog_out(0,0.4)
  	if (Flowability == "LOW"):
  		movel(end_rel_tilted_level2, a=0.03, v=0.1)
  		sleep(0.5)
  		movel(move_inside_spill, a=0.05, v=0.2)
  	  	movel(pose_trans(move_inside_spill, p[0,0,0,0,0,2.0]), a=0.05, v=0.2)
  		#movel(tilted_pose_in_base2, a=0.05, v=0.2)
  	else:
  	    movel(pose_trans(move_inside_spill, p[0,0,0,0,0,2.0]), a=0.05, v=0.2)
  	    movel(move_inside_spill, a=0.05, v=0.2)
  	end
  	set_analog_out(0,0.0)
  	movel(lifted_pose, a=0.5, v=0.5)
  	tilt_to_home()
  	set_tcp(tcp_default)
  end

  def center_pose():
  	global p_translated = container_place
  	#global p_translated = pots_axis_temp

  	#cx = p_translated[0]
  	#cy = p_translated[1]
  	#cz = p_translated[2]

  	global p_center_vertical_temp = pose_trans(p_translated, p[0,0,0, deg2rad(90), 0, 0])
  	cx = p_center_vertical_temp[0]
  	cy = p_center_vertical_temp[1]
  	cz = p_center_vertical_temp[2]
  	rx = p_center_vertical_temp[3]
  	ry = p_center_vertical_temp[4]
  	rz = p_center_vertical_temp[5]

  	global p_center_vertical_temp = p[cx,cy,cz, 0, 0, rz]
  	trans_rel = p[0,0,-pick_2_base+H,0,0,0]
  	global p_center_vertical =  pose_trans(p_center_vertical_temp, trans_rel)
  	return p_center_vertical
  end

  def updated_center_pose(p_center_vertical, angle_deg):
  	hinge_pose = pose_trans(p_center_vertical, p[0,0,-hinge_2_base-gear_2_holder-H ,0,0,0])
  	local_rel = pose_trans(pose_inv(hinge_pose), p_center_vertical)

  	rot_tilt = p[0,0,0, -deg2rad(angle_deg),0,0]
  	local_rel_tilted = pose_trans(rot_tilt, local_rel)

  	global p_center = pose_trans(hinge_pose, local_rel_tilted)
  	return p_center
  end

  def scoop_powder(p_center):
  	vibration_voltage = 0.4
  	global scoop_radius_default = 0.0

  	scoop_radius_default = mouth_d /2 - spatula_depth - wall_thickness
  	scoop_safe_entry_pose = pose_trans(p_center, p[-TCP_2_tip_x,0,spatula_len+0.05,0,0,0])
  	scoop_entry_pose = pose_trans(p_center, p[-TCP_2_tip_x,0,spatula_len,0,0,0])

  	movel(scoop_safe_entry_pose, a=0.1, v=0.25)
  	movel(scoop_entry_pose, a=0.1, v=0.25)

  	scoop_start_rel_int = p[0, 0, -mouth_sh , 0, 0, 0]
  	scoop_start_pose_int = pose_trans(scoop_entry_pose, scoop_start_rel_int)


  	#local ry_deg = map_tilt_to_ry_deg(angle_deg,level)
  	#local ry_result = map_tilt_to_ry_deg(angle_deg,level)

  	#global scoop_depth = compute_scoop_depth(level,weight_value, target_g)

  	global ry = deg2rad(90-angle_deg)

  	#global ry_safe = ry_result[0]
  	#global ry = deg2rad(ry_result[1])

  	if (spatula_mid < powder_height):

  		global total_depth = mouth_sh + scoop_depth + spatula_mid
  		global total_depth = clamp(total_depth, 0, H - spatula_mid)

  		safe_scoop_pivot = (mouth_d  - spatula_depth-wall_thickness)/(total_depth)
  		global ry_safe = asin(safe_scoop_pivot)

  		scoop_start_rel = p[scoop_radius_default, 0, -total_depth, 0, 0, 0]

  		rot_mid = p[0, 0, 0, 0, 0, 0.785]
  		rot_end = p[0, 0, 0, 0, 0, 1.5708]

  		scoop_via_rel = pose_trans(rot_mid, scoop_start_rel)
  		scoop_end_rel = pose_trans(rot_end, scoop_start_rel)

  		scoop_start_pose = pose_trans(scoop_entry_pose, scoop_start_rel)
  		scoop_via_pose = pose_trans(scoop_entry_pose, scoop_via_rel)
  		scoop_end_pose = pose_trans(scoop_entry_pose, scoop_end_rel)


  			if (Flowability == "LOW" and level <= 50):
  				movel(pose_trans(scoop_start_pose_int,p[0,0,0,0,0,-1.5708]), a=0.1, v=0.25)
  				local spatula_base = pose_trans(scoop_entry_pose, p[0, 0, -H+wall_thickness, 0, 0, 0])
  				local scrape_pivot = pose_trans(scoop_entry_pose, p[0,0, -spatula_len,0,0,0])

  				global sticky_in_angle = -atan((cent_edge/2-spatula_depth)/H)
  				spatula_tilt_rel = pose_trans(pose_inv(scrape_pivot), spatula_base)

  				spatula_tilt = pose_trans(spatula_tilt_rel, p[0, 0, 0, 0, sticky_in_angle, 0])
  				global tilted_pose = pose_trans(scrape_pivot, p[0,0,0,spatula_tilt[3],spatula_tilt[4], spatula_tilt[5]])

  				global tilted_pose = pose_trans(tilted_pose, p[0,0,spatula_len-H+wall_thickness,0,0,0])
  				global rotate_90=pose_trans(tilted_pose,p[0,0,0,0,0,-1.5708])
  				movel(rotate_90,a=0.1, v=0.25)
  				CW_full_Rotate()
  				movel(scoop_start_pose, a=0.1, v=0.25)
  			else:
  				movel(scoop_start_pose_int, a=0.1, v=0.25)
  				movel(scoop_start_pose, a=0.1, v=0.25)
  				CW_full_Rotate()
  			end

  		movec(scoop_via_pose, scoop_end_pose, a=0.05, v=0.04)
  		#sleep(1.0)

  		# safe_retention
  		local pivot_pose = pose_trans(scoop_end_pose, p[0,0,total_depth-spatula_len,0,0,0])
  		local end_rel = pose_trans(pose_inv(pivot_pose), scoop_end_pose)
  		local end_rel_tilted = pose_trans(end_rel, p[0, 0, 0, 0, ry_safe-deg2rad(spatula_ry), 0])
  		local tilted_pose_in_base = pose_trans(pivot_pose, p[0,0,0,end_rel_tilted[3],end_rel_tilted[4], end_rel_tilted[5]])
  		local tilted_pose_in_base = pose_trans(tilted_pose_in_base, p[0, 0, spatula_len-total_depth, 0, 0, 0])
  		# sptula pivoted around the container rim of the mouth at ry_safe
  		movel(tilted_pose_in_base, a=0.03, v=0.1)

  		global safe_x = sin(ry_safe)*(total_depth-mouth_sh - (mouth_d - spatula_depth)*tan(ry_safe/2))
  		global safe_z = cos(ry_safe)*(total_depth-mouth_sh - (mouth_d - spatula_depth)*tan(ry_safe/2))

  		local safe_up = pose_trans(tilted_pose_in_base, p[-safe_x,0,safe_z,0,0,0])
  		movel(safe_up, a=0.03, v=0.1)

  		# full exit
  		local pivot_pose2 = pose_trans(scoop_entry_pose, p[0,0,-spatula_len,0,0,0])
  		local end_rel2 = pose_trans(pose_inv(pivot_pose2), tilted_pose_in_base)
  		#popup("is the spatula crashing front? ", blocking = True)
  		local end_rel_tilted2 = pose_trans(end_rel2, p[0, 0, 0, 0, ry-ry_safe-deg2rad(spatula_ry), 0])

  	else : # emptying logic
  		#CCW_full_Rotate()

  		spatula_base = pose_trans(scoop_entry_pose, p[0, 0, -H+wall_thickness, 0, 0, 0])
  		local pivot_pose2 = pose_trans(scoop_entry_pose, p[0,0,-spatula_len,0,0,0])
  		# tilt inwards
  		global in_angle = -atan((cent_edge/2-spatula_depth)/H)
  		spatula_tilt_rel = pose_trans(pose_inv(pivot_pose2), spatula_base)

  		spatula_tilt = pose_trans(spatula_tilt_rel, p[0, 0, 0, -in_angle, 0, 0])
  		global tilted_pose = pose_trans(pivot_pose2, p[0,0,0,spatula_tilt[3],spatula_tilt[4], spatula_tilt[5]])

  		global tilted_pose = pose_trans(tilted_pose, p[0,0,spatula_len-H+wall_thickness,0,0,0])

  		movel(tilted_pose,a=0.1, v=0.25)
  		CW_full_Rotate()
  		sleep(1)
  		rotate90=pose_trans(tilted_pose,p[0,0,0,0,0,1.5708])

  		#sleep(1)
  		#Rotate()
  		#sleep(0.2)
  		movel(rotate90, a=0.1, v=0.1)
  		#popup("is the spatula crashing front? ", blocking = True)
  		movel(pose_trans(scoop_start_pose_int,p[0,0,0,0,0,1.5708]), a=0.03, v=0.1)
  		# full exit
  		#local pivot_pose2 = pose_trans(scoop_entry_pose, p[0,0,-spatula_len,0,0,0])
  		local end_rel2 = pose_trans(pose_inv(scoop_entry_pose), rotate90)
  		local end_rel_tilted2 = pose_trans(end_rel2, p[0, 0, 0, 0, ry-in_angle-deg2rad(spatula_ry), 0])
  	end

  	# exit flat spoon
  	global tilted_pose_in_base2 = pose_trans(pivot_pose2, p[0,0,0,end_rel_tilted2[3],end_rel_tilted2[4], end_rel_tilted2[5]])
  	global tilted_pose_in_base2 = pose_trans(tilted_pose_in_base2, p[0, 0, spatula_len-spatula_mid, 0, 0, 0])
  	# spaula exited at center of the mouth at ry
  	movel(tilted_pose_in_base2, a=0.03, v=0.1)

  	if(spatula == "spatula_S"):
  		if(level>=80):
  			global z_ratio = 0.0
  		elif(level == 0.0):
  			global z_ratio = 1.0
  		else:
  			global z_ratio = (80-level)/80
  		end
  		z_offset = 4*spatula_mid*z_ratio
  	elif(spatula == "spatula_flat_S"):
  		if(level>=50):
  			global z_ratio = 0.0
  		elif(level == 0.0):
  			global z_ratio = 1.0
  		else:
  			global z_ratio = (50-level)/50
  		end
  		z_offset = 4*spatula_mid*z_ratio
  	else:
  	    z_offset = 0.0
  	end

  	global move_inside_spill = pose_trans(tilted_pose_in_base2, p[0,0,-z_offset,0,0,0])
  	movel(move_inside_spill, a=0.03, v=0.1)

  	if(scoop_status== "normal"):
  		vib_thread=True
  		if (spatula=="spatula_S"):
  			vibration_3()
  			local ry_level = deg2rad(5)
  		elif(spatula=="spatula_flat_S" or spatula=="spatula_flat_M"):
  			vibration_3()
  			local ry_level = deg2rad(5)
  		else:
  			set_analog_out(0,0.4)
  			local ry_level = deg2rad(15)
  		end

  		# remove excess
  		local pivot_pose_level = pose_trans(move_inside_spill, p[0,0,-spatula_len,0,0,0])
  		local end_rel_level = pose_trans(pose_inv(pivot_pose_level), move_inside_spill)
  		local end_rel_tilted_level = pose_trans(end_rel_level, p[0, 0, 0, 0, -ry_level, 0])
  		global end_rel_tilted_level2 = pose_trans(pivot_pose_level, p[0, 0, 0,end_rel_tilted_level[3],end_rel_tilted_level[4], end_rel_tilted_level[5]])
  		global end_rel_tilted_level2 = pose_trans(end_rel_tilted_level2, p[0,0,spatula_len,0,0,0])
  		movel(end_rel_tilted_level2, a=0.03, v=0.1)

  		if (spatula == "spatula_flat_S" or spatula == "spatula_flat_M"):
  			vib_thread=False
  			set_analog_out(0, 0.0)
  		end
  	else:
  		set_analog_out(0, 0.0)
  	end
  	movel(tilted_pose_in_base2, a=0.03, v=0.1)
  	set_analog_out(0, 0.0)
  	vib_thread=False
  	global lifted_pose = pose_trans(tilted_pose_in_base2, p[-0.04,0,0.04,0,0,0]) # safety distance away from the container

  	movel(lifted_pose, a=0.03, v=0.1)
  	tilt_to_home()
  end

  def auto_tilt_and_scoop(W_now, target_weight, weight_value):
  	set_tcp(tcp_dosing)
  	#global level = compute_level_percent(W_now, weight_value)

  	global spatula = select_spatula(Flowability, level, diff, bulk_density, mouth_d )
  	textmsg("deb 4 = ", spatula)
  	global target_g = get_scoop_weight(spatula, bulk_density)
  	textmsg("deb 5 = ", target_g)

  	global scoop_depth = compute_scoop_depth(level, weight_value, target_g)
    	textmsg("deb 6 = ", scoop_depth)
  	tilt(level)

  	scoop_powder(p_center)

  	#textmsg("deb 7 - sucess")
   	set_tcp(tcp_default)
  end
  $ 21 "Script: Weight_scale_socket_s.script"
  global s_depth = 0
  global s_length =0
  global s_volume = 0
  global ry_theta  = 0

  def get_weight():
  	socket_open(SERVER_IP,SERVER_PORT)
  	#sleep(0.2)
  	textmsg("socket opened successfully!")
  	socket_send_string("GET_WEIGHT")
  	#sleep(0.2)
  	sync()
  	receiveFromServ = socket_read_ascii_float(1)
  	#sleep(1)
  	while (receiveFromServ[0] < 1):
  		receiveFromServ = socket_read_ascii_float(1)
  		sleep(0.01)
  	end
  	textmsg("Received weight:", receiveFromServ[1])
  	#sleep(0.2)
  	socket_close()
  	#sleep(0.2)
  	return receiveFromServ[1]
  end

  def tare_scale():
  	socket_open(SERVER_IP,SERVER_PORT)
  	socket_send_string("TARE")
  	sleep(2)
  	socket_close()
  end

  def zero_scale():
  	socket_open(SERVER_IP,SERVER_PORT)
  	socket_send_string("ZERO")
  	sleep(0.5)
  	socket_close()
  end

  def log_weight():
  	socket_open(SERVER_IP,SERVER_PORT)
  	socket_send_string("LOG_WEIGHT")
  	sleep(0.5)
  	socket_close()
  end

  def send_target_info():
  	socket_open(SERVER_IP,SERVER_PORT)
  	socket_send_string("SET_TARGET:" + to_str(target_weight))
  	sleep(0.2)
  	socket_close()
  end
  def send_powder_info():
  	socket_open(SERVER_IP,SERVER_PORT)
  	socket_send_string("SET_POWDER:" + Pow_name)
  	sleep(0.2)
  	socket_close()
  end
  def send_spatula_info():
  	socket_open(SERVER_IP,SERVER_PORT)
  	socket_send_string("SET_SPATULA:" + spatula)
  	#sleep(1)

  	#local fl = socket_read_ascii_float(4)

    	#global s_depth = fl[1]
    	#global s_length = fl[2]
   	#global s_volume = fl[3]
   	#global ry_theta  = fl[4]
  	sleep(0.2)
  	socket_close()
  end

  def send_level_info():
  	socket_open(SERVER_IP,SERVER_PORT)
  	socket_send_string("SET_LEVEL:" + to_str(level))
  	sleep(0.2)
  	socket_close()
  end

  def get_cont_weight():
    socket_open(SERVER_IP, SERVER_PORT)
    #rq_open_and_wait()
    cmd = "GET_CONT_WEIGHT"
    socket_send_string(cmd)
    sync()
    sleep(0.5)
    receiveFromSer = socket_read_ascii_float(1)
    socket_close()
    return receiveFromSer[1]
  end

  $ 22 "Script: swab_sampling.script"
  global swab_poses=make_list(0,0,6)
  global pose_list_hor=make_list(0,0,420)
  global pose_list_ver=make_list(0,0,420)
  global cntd=False
  global trgt_waypts=make_list(0,0,6)
  global new_z=0
  global first_pts=make_list(0,0,15)
  global temp_pose_force=p[0,0,0,0,0,0]
  global delta_rx=0
  global new_dz=0
  global server_msg=""
  global delta_x=0
  global delta_y=0


  def connect2server():
  	IP="192.168.12.139"
  	port=3002
  	while(cntd==False):
  		cntd=socket_open(IP,port)
  		if(cntd==True):
  			textmsg("Connected to server")
  		end
  	end
  	socket_send_string("SCAN_TARGET")
  end


  def get_hor_pose_from_server():

  	IP="192.168.12.139"
  	port=3002
  	if(cntd==True):
  		textmsg("Connected to server")
  	end
  	while(cntd==False):
  		cntd=socket_open(IP,port)
  		if(cntd==True):
  			textmsg("Connected to server")
  		end
  		sleep(0.2)
  	end
  	socket_send_string("GET_POSE_HOR")
  	idx=socket_read_ascii_float(1,timeout=-1)
  	textmsg("Index from server=",idx[1])
  	itn_i=0
  	while(itn_i<idx[1]):
  		msg=socket_read_ascii_float(6,timeout=-1)
  		i=1
  		while(i<7):
  			swab_poses.append(msg[i])
  			i=i+1
  		end
  		pose_list_hor.extend(swab_poses)
  		swab_poses.clear()
  		socket_send_string("OK")
  		itn_i=itn_i+1
  	end
  	socket_read_line(timeout=-1)
  	if(cntd==True):
  		cntd=False
  		socket_close()
  	end
  	#textmsg("server msg",swab_poses)
  	textmsg("pose list",pose_list_hor)
  end


  def get_ver_pose_from_server():
  	IP="192.168.12.139"
  	port=3002
  	if(cntd==True):
  		textmsg("Connected to server")
  	end
  	while(cntd==False):
  		cntd=socket_open(IP,port)
  		if(cntd==True):
  			textmsg("Connected to server")
  		end
  		sleep(0.2)
  	end
  	socket_send_string("GET_POSE_VER")
  	idx=socket_read_ascii_float(1,timeout=-1)
  	textmsg("Index from server=",idx[1])
  	itn_i=0
  	while(itn_i<idx[1]):
  		msg=socket_read_ascii_float(6,timeout=-1)
  		i=1
  		while(i<7):
  			swab_poses.append(msg[i])
  			i=i+1
  		end
  		pose_list_ver.extend(swab_poses)
  		swab_poses.clear()
  		socket_send_string("OK")
  		itn_i=itn_i+1
  	end
  	socket_read_line(timeout=-1)
  	if(cntd==True):
  		cntd=False
  		socket_close()
  	end
  	#textmsg("server msg",swab_poses)
  	textmsg("pose list",pose_list_ver)
  end


  def move_to_first_point(code):
  	first_pts.clear()
  	k=0
  	i=1
  	l=1
  	blend_r=0
  	while(i<3):
  		j=1
  		while(j<=6):
  			k=l-1
  			if(code==1):
  				first_pts.append(pose_list_hor[k])
  			elif(code==2):
  				first_pts.append(pose_list_ver[k])
  			end
  			j=j+1
  			l=l+1
  		end
  		i=i+1
  	end
  	movel(p[first_pts[0]-delta_y,first_pts[1]+delta_x,first_pts[2],first_pts[3],first_pts[4],first_pts[5]],a=0.5,v=0.05,r=blend_r)
  	sleep(2)
  	zero_ftsensor()
  	sleep(2)
  	tcp_f=get_tcp_force()
  	textmsg("Force after zeroing:",tcp_f)
  	ftmode=True
  	while(ftmode==True):
  		tcp_f=get_tcp_force()
  		if tcp_f[2]<0.7:
  			speedl([0,0,-0.001,0,0,0],0.05,t=0.5)
  		else:
  			stopl(3)
  			new_p=get_actual_tcp_pose()
  			new_z=new_p[2]-first_pts[2]
  			ftmode=False
  		end
  		sleep(0.2)
  	end
  	movel(p[first_pts[6]-delta_y,first_pts[7]+delta_x,first_pts[8]+new_z,first_pts[9],first_pts[10],first_pts[11]],a=0.5,v=0.05,r=blend_r)
  	curr_tcp=get_actual_tcp_pose()
  	textmsg("Current TCP",curr_tcp)
  	#tcp_str=to_string(curr_tcp)
  	popup("Tcp change",blocking=True)
  	#temp_pose_force=p[first_pts[0],first_pts[1],first_pts[2],first_pts[3],first_pts[4],first_pts[5]]
  	temp_pt=first_pts[2]
  	first_pts.clear()
  	zero_ftsensor()
  	sleep(2)
  	tcp_f=get_tcp_force()
  	textmsg("Force after zeroing:",tcp_f)
  	ftmode=True
  	#ftmode=False
  	while(ftmode==True):
  		tcp_f=get_tcp_force()
  		textmsg("Force",tcp_f)
  		if tcp_f[2]<2.5:
  			speedl([0,0,-0.005,0,0,0],0.05,t=0.5)
  		else:
  			stopl(3)
  			new_p=get_actual_tcp_pose()
  			new_dz=new_p[2]-temp_pt
  			ftmode=False
  			textmsg("DZ=",new_dz)
  		end
  		sleep(0.2)
  	end
  	IP="192.168.12.139"
  	port=3002
  	if(cntd==True):
  		textmsg("Connected to server")
  	end
  	while(cntd==False):
  		cntd=socket_open(IP,port)
  		if(cntd==True):
  			textmsg("Connected to server")
  		end
  		sleep(0.2)
  	end
  	socket_send_string("POSE")
  	socket_send_string(str_cat("",curr_tcp))
  	if(cntd==True):
  		cntd=False
  		socket_close()
  	end

  end

  def follow_swab_trajectory_hor():
  	idx=pose_list_hor.length()
  	textmsg("idx",idx)
  	idx=idx/6
  	k=0
  	i=3
  	l=13
  	delta_z=0.035
  	zero_ftsensor()
  	sleep(1)
  	#tcp_f=get_tcp_force()
  	#textmsg("Force at tip:",tcp_f)
  	force_mode(temp_pose_force,[0,0,1,0,0,0],[0,0,0.3,0,0,0],2,[0.005,0.005,0.05,0.01,0.01,0.01])
  	while(i<=idx):
  		j=1
  		while(j<=6):
  			k=l-1
  			trgt_waypts.append(pose_list_hor[k])
  			j=j+1
  			l=l+1
  		end
  		if(i<3):
  			delta_rx=0
  			delta_z=0
  			blend_r=0
  		elif((i-1)%5==0):
  			blend_r=0
  			delta_z=0.043
  			#delta_rx=0.104
  			delta_rx=0.3
  		else:
  			blend_r=0.002
  			delta_z=0.043
  			#delta_rx=0.104
  			delta_rx=0.3
  		end
  		if(i==1):
  			delta_z=0.005
  			trgt_waypts[2]=trgt_waypts[2]+delta_z
  		movel(p[trgt_waypts[0],trgt_waypts[1],trgt_waypts[2],trgt_waypts[3],trgt_waypts[4],trgt_waypts[5]],a=0.5,v=0.05,r=blend_r)
  			zero_ftsensor()
  			sleep(1)
  			ftmode=True
  			while(ftmode==True):
  				tcp_f=get_tcp_force()
  				if tcp_f[2]<0.7:
  					speedl([0,0,-0.001,0,0,0],0.5,t=0.5)
  				else:
  					stopl(3)
  					new_p=get_actual_tcp_pose()
  					new_z=new_p[2]-trgt_waypts[2]
  					textmsg("Force at tip:",tcp_f)
  					ftmode=False
  				end
  				sleep(0.2)
  			end
  		else:

  			delta_z=0
  			trgt_waypts[2]=trgt_waypts[2]+new_z+delta_z+new_dz
  			trgt_waypts[3]=trgt_waypts[3]-delta_rx
  		movel(p[trgt_waypts[0],trgt_waypts[1],trgt_waypts[2],trgt_waypts[3],trgt_waypts[4],trgt_waypts[5]],a=0.5,v=0.01,r=blend_r)
  			tcp_f=get_tcp_force()
  			#tcp_f=get_tcp_force_tool()
  			textmsg("Force at tip:",tcp_f)
  		end
  		textmsg("Target Waypoints",trgt_waypts)
  		trgt_waypts.clear()
  		i=i+1
  	end
  	end_force_mode()
  	pose_list_hor.clear()
  end

  def follow_swab_trajectory(code):
  	dy=0.036
  	pose_list_temp=make_list(0,0,420)
  	if(code==1):
  		pose_list_temp=pose_list_hor
  		delta_x=0
  		delta_y=0
  	elif(code==2):
  		pose_list_temp=pose_list_ver
  	end
  	idx=pose_list_temp.length()
  	textmsg("idx",idx)
  	idx=idx/6
  	k=0
  	i=3
  	l=13

  	zero_ftsensor()
  	sleep(2)
  	IP="192.168.12.139"
  	port=3002
  	if(cntd==True):
  		textmsg("Connected to server")
  	end
  	while(cntd==False):
  		cntd=socket_open(IP,port)
  		if(cntd==True):
  			textmsg("Connected to server")
  		end
  		sleep(0.2)
  	end
  	#force_mode(temp_pose_force,[0,0,1,0,0,0],[0,0,1,0,0,0],2,[0.001,0.001,0.01,0.01,0.01,0.01])
  	while(i<=idx):
  		socket_send_string("PLOT")
  		j=1
  		while(j<=6):
  			k=l-1
  			trgt_waypts.append(pose_list_temp[k])
  			j=j+1
  			l=l+1
  		end
  		if(i<3):
  			delta_rx=0
  			delta_z=0
  			blend_r=0
  		elif((i-1)%5==0):
  			blend_r=0
  			#delta_z=0.043
  			#delta_rx=0.104
  			delta_rx=0.3
  		else:
  			blend_r=0.002
  			#delta_z=0.043
  			#delta_rx=0.104
  			delta_rx=0.3
  		end
  		delta_z=0
  		if(i==3):
  			temp=get_actual_tcp_pose()
  			delta_y=temp[1]-trgt_waypts[1]
  			delta_x=temp[0]-trgt_waypts[0]
  		end
  		#textmsg("delta Y:",delta_y)
  		#textmsg("delta X:",delta_x)
  		delta_x=0
  		delta_y=0
  		trgt_waypts[0]=trgt_waypts[0]+delta_x
  		trgt_waypts[1]=trgt_waypts[1]+delta_y
  		trgt_waypts[2]=trgt_waypts[2]+new_dz 		#new_z
  		trgt_pose=pose_trans(p[trgt_waypts[0],trgt_waypts[1],trgt_waypts[2],trgt_waypts[3],trgt_waypts[4],trgt_waypts[5]],p[0,0,0,0,0,0])
  		movel(trgt_pose,a=0.5,v=0.005,r=blend_r)
  		tcp_f=get_tcp_force()
  		#textmsg("Force at tip:",tcp_f)
  		#textmsg("Target Waypoints",trgt_waypts)
  		trgt_waypts.clear()
  		i=i+1
  	end
  	#end_force_mode()
  	socket_send_string("PLOT DONE")
  	if(cntd==True):
  		cntd=False
  		socket_close()
  	end
  	#speedl([0,0,0.05,0,0,0],0.05,t=0.5)
  	pose_list_temp.clear()
  	if(code==2):
  		delta_x=0
  		delta_y=0
  	end
  end


  def follow_swab_trajectory_ver():
  	idx=pose_list_ver.length()
  	textmsg("idx",idx)
  	idx=idx/6
  	k=0
  	i=1
  	l=1
  	while(i<=idx):
  		j=1
  		while(j<=6):
  			k=l-1
  			trgt_waypts.append(pose_list_ver[k])
  			j=j+1
  			l=l+1
  		end
  		movel(p[trgt_waypts[0],trgt_waypts[1],trgt_waypts[2],trgt_waypts[3],trgt_waypts[4],trgt_waypts[5]],a=0.5,v=0.2)
  		textmsg("Target Waypoints",trgt_waypts)
  		trgt_waypts.clear()
  		i=i+1
  	end
  	pose_list_ver.clear()
  end


  def wait_acknowledge():
  	pose_list_hor.clear()
  	pose_list_ver.clear()
  	IP="192.168.12.139"
  	port=3002
  	if(cntd==True):
  		textmsg("already Connected to server")
  	end
  	while(cntd==False):
  		cntd=socket_open(IP,port)
  		if(cntd==True):
  			textmsg("Connected to server")
  		end
  		sleep(0.2)
  	end
  	serv_msg=socket_read_line(timeout=-1)
  	textmsg("Server Message",serv_msg)

  	if(cntd==True):
  		cntd=False
  		socket_close()
  	end
  	return serv_msg

  end

  def disconnectfromserver():
  	delta_x=0
  	delta_y=0
  	socket_close()
  end

  def swab_break():
  	curr_tcp=get_actual_tcp_pose()
  	brk_pt=pose_add(curr_tcp,p[0,0,0.04,0,0,0])
  	popup("tcp_changed to breaking point",blocking=True)
  	movel(pose_trans(brk_pt,p[0,0,0,0,1.3,0]),a=0.5,v=0.005)
  	#movel(p[brk_pt[0],brk_pt[1],brk_pt[02],brk_pt[3],brk_pt[4]+1.57,brk_pt[5]],a=0.5,v=0.005)
  end

  #Helper Function

  def get_tcp_force_tool():
  	force_torque= get_tcp_force()
  	force_B=p[force_torque[0],force_torque[1],force_torque[2],0,0,0]
  	torque_B=p[force_torque[3],force_torque[4],force_torque[5],0,0,0]
  	tcp=temp_pose_force
  	rotation_BT=p[0,0,0,tcp[3],tcp[4],tcp[5]]
  	force_T= pose_trans(pose_inv(rotation_BT),force_B)
  	torque_T=pose_trans(pose_inv(rotation_BT),torque_B)
  	force_torque_T=p[force_T[0],force_T[1],force_T[2],torque_T[0],torque_T[1],torque_T[2]]
  	return force_torque_T
  end




  $ 23 "BeforeStarts"
  $ 24 "uLM"
  $ 25 "CMD_Stop≔ False "
  global CMD_Stop=  False
  $ 26 "CMD_Abort≔ False "
  global CMD_Abort=  False
  $ 27 "CMD_Clear≔ False "
  global CMD_Clear=  False
  $ 28 "STATE≔1"
  global STATE=1
  $ 29 "STATE_Info≔''"
  global STATE_Info=""
  $ 30 "ARM_Referenced≔ False "
  global ARM_Referenced=  False
  $ 31 "zero_ftsensor()"
  zero_ftsensor()
  $ 32 "poses init"
  $ 33 "PSE_A≔p[0,0,0,0,0,0]"
  global PSE_A=p[0,0,0,0,0,0]
  $ 34 "PSE_A_H≔p[0,0,0,0,0,0]"
  global PSE_A_H=p[0,0,0,0,0,0]
  $ 35 "PSE_R≔p[0,0,0,0,0,0]"
  global PSE_R=p[0,0,0,0,0,0]
  $ 36 "PSE_R_H≔p[0,0,0,0,0,0]"
  global PSE_R_H=p[0,0,0,0,0,0]
  $ 37 "PSE_T≔p[0,0,0,0,0,0]"
  global PSE_T=p[0,0,0,0,0,0]
  $ 38 "PSE_T_H≔p[0,0,0,0,0,0]"
  global PSE_T_H=p[0,0,0,0,0,0]
  $ 39 "PSE_C_E≔p[0,0,0,0,0,0]"
  global PSE_C_E=p[0,0,0,0,0,0]
  $ 40 "PSE_C_H≔p[0,0,0,0,0,0]"
  global PSE_C_H=p[0,0,0,0,0,0]
  $ 41 "PSE_C_S≔p[0,0,0,0,0,0]"
  global PSE_C_S=p[0,0,0,0,0,0]
  $ 42 "init_home_by_cartesian_pose(p[0,-0.400,0.300,0,0,0])"
  init_home_by_cartesian_pose(p[0,-0.400,0.300,0,0,0])
  $ 43 "Clearing"
  $ 44 "reset_error()"
  reset_error()
  $ 45 "reset_warning()"
  reset_warning()
  $ 46 "uGo"
  $ 48 "ugo_init( True ,'http://192.168.12.120:10001')"
  ugo_init(  True  ,"http://192.168.12.120:10001")
  $ 49 "ugo_update_outputs()"
  ugo_update_outputs()
  $ 50 "App"
  $ 51 "'ADD APPLICATION SPECIFIC COMMANDS'"
  # 'ADD APPLICATION SPECIFIC COMMANDS'
  $ 52 "Tools"
  $ 53 "OBJ_Picked≔gripper_has_object()"
  global OBJ_Picked=gripper_has_object()
  $ 54 "If OBJ_Picked"
  if (OBJ_Picked):
    # begin: URCap Program Node
    #   Source: Robotiq_Grippers, 3.17.0.105337, Robotiq Inc.
    #   Type: Gripper Activate
    $ 55 "Gripper Activate"

    kill rq_gripper_communication_thread
    rq_gripper_communication_thread_started = False
    rq_close_gripper_socket("1")
    rq_close_gripper_socket("2")
    rq_close_gripper_socket("3")
    rq_close_gripper_socket("4")

    rq_init_comm_if_connected(9, "1")
    rq_init_comm_if_connected(2, "2")
    rq_init_comm_if_connected(3, "3")
    rq_init_comm_if_connected(4, "4")
    rq_print_connected_grippers()
    rq_gripper_communication_thread = run rq_gripper_communication()

    while(not rq_gripper_communication_thread_started):
        sleep(0.008)
    end

    rq_set_max_current_for_all_grippers()

    reset_and_activate = False

    rq_activate_all_grippers(False)
    # end: URCap Program Node
  else:
    $ 56 "Else" "noBreak"
    # begin: URCap Program Node
    #   Source: Robotiq_Grippers, 3.17.0.105337, Robotiq Inc.
    #   Type: Gripper Activate
    $ 57 "Gripper Reset and Activate"

    kill rq_gripper_communication_thread
    rq_gripper_communication_thread_started = False
    rq_close_gripper_socket("1")
    rq_close_gripper_socket("2")
    rq_close_gripper_socket("3")
    rq_close_gripper_socket("4")

    rq_init_comm_if_connected(9, "1")
    rq_init_comm_if_connected(2, "2")
    rq_init_comm_if_connected(3, "3")
    rq_init_comm_if_connected(4, "4")
    rq_print_connected_grippers()
    rq_gripper_communication_thread = run rq_gripper_communication()

    while(not rq_gripper_communication_thread_started):
        sleep(0.008)
    end

    rq_set_max_current_for_all_grippers()

    reset_and_activate = True

